// TIA Portal V20 export
// export: Created 2026-10-20T18:54:23.1624492Z, ExportSetting None, DisplayName Totally Integrated Automation Portal, DisplayVersion V20 Update 6, DisplayName TIA Portal Openness, DisplayVersion V20 Update 6, DisplayName TIA Portal Version Control Interface, DisplayVersion V20 Update 6, DisplayName SINAMICS Startdrive Advanced, DisplayVersion V20 SP1, DisplayName SINAMICS Startdrive G130, G150, S120, S150, SINAMICS MV, G220, S200, S210, DisplayVersion V20 SP1, DisplayName SINAMICS Startdrive G110M, G120, G120C, G120D, G120P, G115D, DisplayVersion V20 SP1, DisplayName STEP 7 Professional, DisplayVersion V20 Update 6, DisplayName STEP 7 Safety, DisplayVersion V20 Update 2, DisplayName WinCC Basic/Comfort/Advanced, DisplayVersion V20 Update 6, DisplayName WinCC Unified, DisplayVersion V20 Update 6
VAR_GLOBAL   // PLC tag table "CNV_HMI_IO"
   "HMI_CNV_SftyPinDown(1)" AT %M2.3 : Bool;
   HMI_CNV_SftyPinDown AT %M1.1 : Bool;
   HMI_CNV_Sdetect1 AT %M0.6 : Bool;
   "HMI_CNV_SftyPinUp(1)" AT %M2.2 : Bool;
   HMI_CNV_Sdetect2 AT %M0.7 : Bool;
   HMI_CNV_SftyPinUp AT %M1.0 : Bool;
   "HMI_CNV_Sdetect1(1)" AT %M2.0 : Bool;
   "HMI_CNV_Sdetect2(1)" AT %M2.1 : Bool;
   "HMI_CNV_Rpd2(1)" AT %M1.7 : Bool;
   HMI_CNV_Lpd2 AT %M0.2 : Bool;
   "HMI_CNV_Rpd1(1)" AT %M1.6 : Bool;
   "HMI_CNV_Lpd2(1)" AT %M1.4 : Bool;
   "HMI_CNV_Lpd1(1)" AT %M1.3 : Bool;
   HMI_CNV_Rpd1 AT %M0.4 : Bool;
   HMI_CNV_Lpd1 AT %M5.6 : Bool;
   HMI_CNV_Rpd2 AT %M0.5 : Bool;
   "HMI_CNV_Right(1)" AT %M1.5 : Bool;
   HMI_CNV_Right AT %M0.3 : Bool;
   HMI_CNV_Left AT %M0.0 : Bool;
   "HMI_CNV_Left(1)" AT %M1.2 : Bool;
   HMI_Light_Guard AT %M61.4 : Bool;
END_VAR
